INTERFACE I_DigitalOut

METHOD SwitchOn
END_METHOD

METHOD SwitchOff
END_METHOD

PROPERTY IsOn : BOOL
GET
END_GET
END_PROPERTY

END_INTERFACE

(* stored: Version 1.1.0.1, ProductVersion 3.1.4026.12
   Itf I_DigitalOut: Id {2fec7f26-66ea-510e-8e2c-720bc689c950}
   Method SwitchOn: Id {2c722ea5-f2c4-50e0-aeb5-4edd0b0fb292}
   Method SwitchOff: Id {faa4dbff-6904-5b2d-b91a-18fec5c4fb79}
   Property IsOn: Id {f8359847-95c8-59d4-871a-3479d5cf994e}
   Get Get: Id {67236b3f-0699-5e1a-945b-2d4e38a64259} *)
